// Mitsubishi GX Works2 project: SEMICON_SORTER_ENV   PLC: FX3U/FX3UC

PROGRAM MAIN
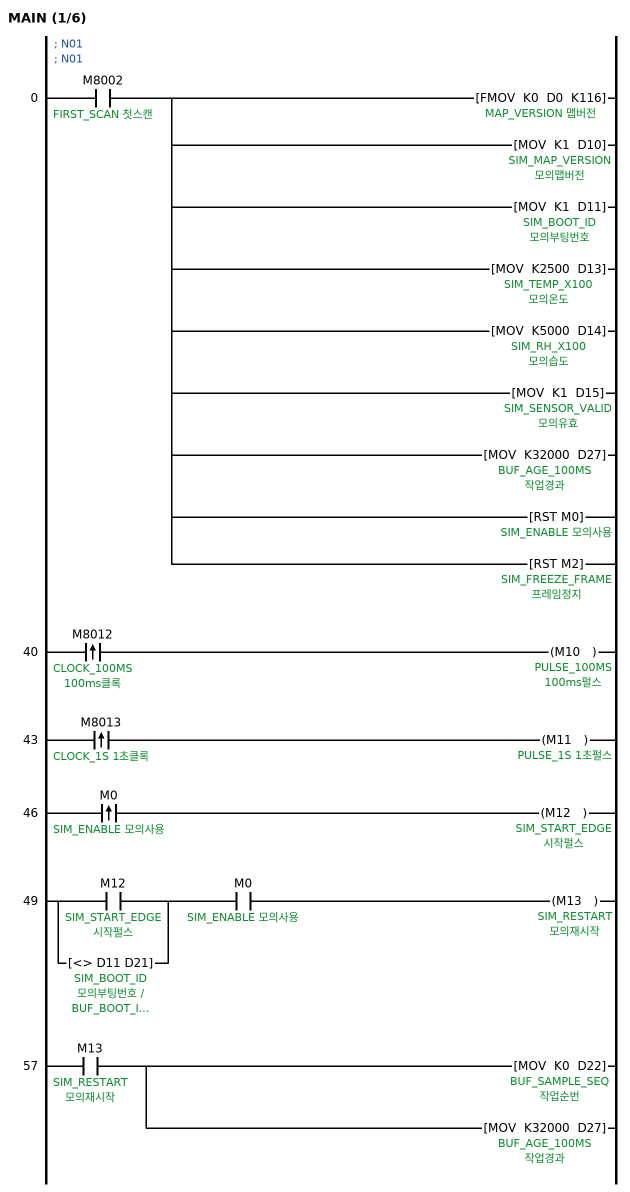
; 
; N01
; N01
0     LD      M8002  ; FIRST_SCAN 첫스캔
      FMOV    K0 D0 K116  ; MAP_VERSION 맵버전
      MOV     K1 D10  ; SIM_MAP_VERSION 모의맵버전
      MOV     K1 D11  ; SIM_BOOT_ID 모의부팅번호
      MOV     K2500 D13  ; SIM_TEMP_X100 모의온도
      MOV     K5000 D14  ; SIM_RH_X100 모의습도
      MOV     K1 D15  ; SIM_SENSOR_VALID 모의유효
      MOV     K32000 D27  ; BUF_AGE_100MS 작업경과
      RST     M0  ; SIM_ENABLE 모의사용
      RST     M2  ; SIM_FREEZE_FRAME 프레임정지
40    LDP     M8012  ; CLOCK_100MS 100ms클록
      OUT     M10  ; PULSE_100MS 100ms펄스
43    LDP     M8013  ; CLOCK_1S 1초클록
      OUT     M11  ; PULSE_1S 1초펄스
46    LDP     M0  ; SIM_ENABLE 모의사용
      OUT     M12  ; SIM_START_EDGE 시작펄스
49    LD      M12  ; SIM_START_EDGE 시작펄스
      OR<>    D11 D21  ; SIM_BOOT_ID 모의부팅번호 / BUF_BOOT_ID 작업부팅번호
      AND     M0  ; SIM_ENABLE 모의사용
      OUT     M13  ; SIM_RESTART 모의재시작
57    LD      M13  ; SIM_RESTART 모의재시작
      MOV     K0 D22  ; BUF_SAMPLE_SEQ 작업순번
      MOV     K32000 D27
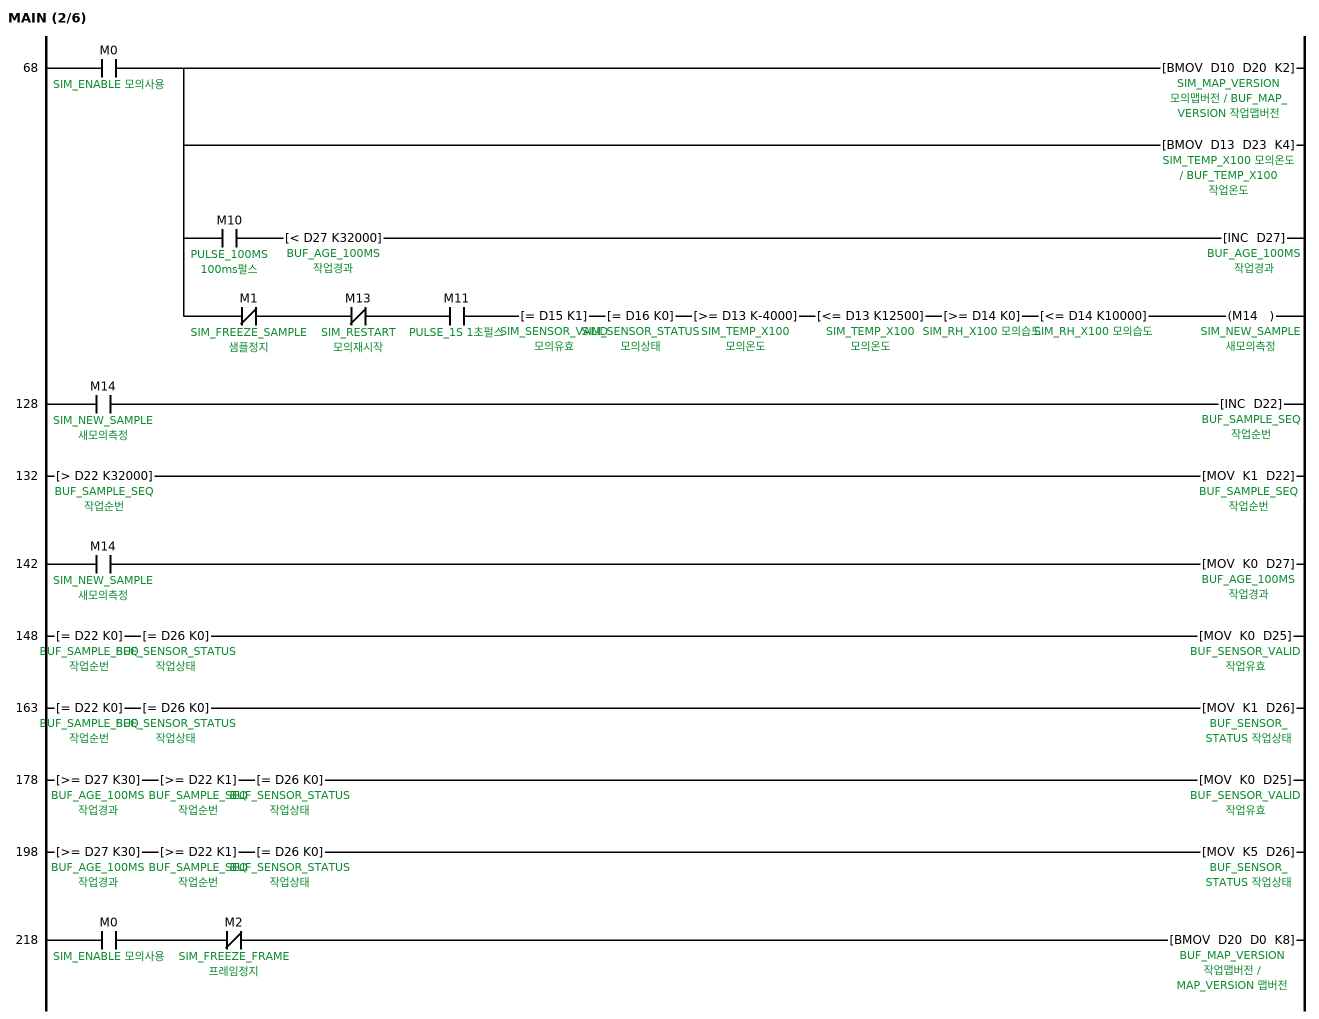
68    LD      M0  ; SIM_ENABLE 모의사용
      BMOV    D10 D20 K2  ; BUF_MAP_VERSION 작업맵버전
      BMOV    D13 D23 K4  ; BUF_TEMP_X100 작업온도
      MPS
      AND     M10  ; PULSE_100MS 100ms펄스
      AND<    D27 K32000  ; BUF_AGE_100MS 작업경과
      INC     D27
      MPP
      ANI     M1  ; SIM_FREEZE_SAMPLE 샘플정지
      ANI     M13  ; SIM_RESTART 모의재시작
      AND     M11  ; PULSE_1S 1초펄스
      AND=    D15 K1  ; SIM_SENSOR_VALID 모의유효
      AND=    D16 K0  ; SIM_SENSOR_STATUS 모의상태
      AND>=   D13 K-4000  ; SIM_TEMP_X100 모의온도
      AND<=   D13 K12500  ; SIM_TEMP_X100 모의온도
      AND>=   D14 K0  ; SIM_RH_X100 모의습도
      AND<=   D14 K10000  ; SIM_RH_X100 모의습도
      OUT     M14  ; SIM_NEW_SAMPLE 새모의측정
128   LD      M14  ; SIM_NEW_SAMPLE 새모의측정
      INC     D22
132   LD>     D22 K32000  ; BUF_SAMPLE_SEQ 작업순번
      MOV     K1 D22
142   LD      M14  ; SIM_NEW_SAMPLE 새모의측정
      MOV     K0 D27
148   LD=     D22 K0  ; BUF_SAMPLE_SEQ 작업순번
      AND=    D26 K0  ; BUF_SENSOR_STATUS 작업상태
      MOV     K0 D25  ; BUF_SENSOR_VALID 작업유효
163   LD=     D22 K0  ; BUF_SAMPLE_SEQ 작업순번
      AND=    D26 K0  ; BUF_SENSOR_STATUS 작업상태
      MOV     K1 D26
178   LD>=    D27 K30  ; BUF_AGE_100MS 작업경과
      AND>=   D22 K1  ; BUF_SAMPLE_SEQ 작업순번
      AND=    D26 K0  ; BUF_SENSOR_STATUS 작업상태
      MOV     K0 D25
198   LD>=    D27 K30  ; BUF_AGE_100MS 작업경과
      AND>=   D22 K1  ; BUF_SAMPLE_SEQ 작업순번
      AND=    D26 K0  ; BUF_SENSOR_STATUS 작업상태
      MOV     K5 D26
218   LD      M0  ; SIM_ENABLE 모의사용
      ANI     M2  ; SIM_FREEZE_FRAME 프레임정지
      BMOV    D20 D0 K8
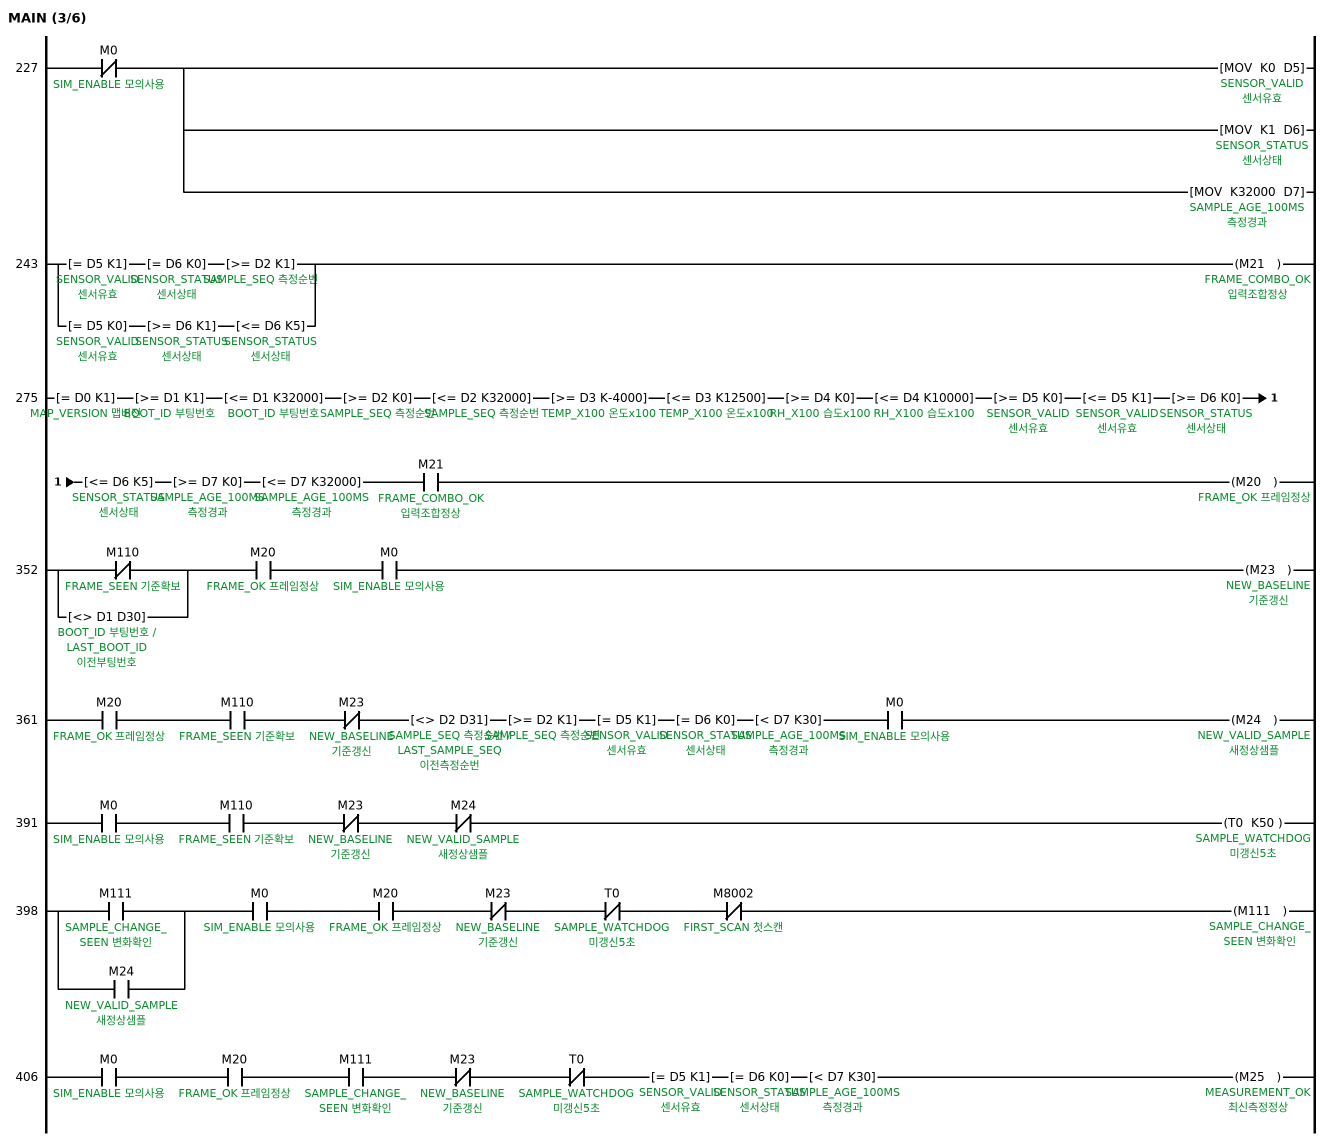
227   LDI     M0  ; SIM_ENABLE 모의사용
      MOV     K0 D5  ; SENSOR_VALID 센서유효
      MOV     K1 D6  ; SENSOR_STATUS 센서상태
      MOV     K32000 D7  ; SAMPLE_AGE_100MS 측정경과
243   LD=     D5 K1  ; SENSOR_VALID 센서유효
      AND=    D6 K0  ; SENSOR_STATUS 센서상태
      AND>=   D2 K1  ; SAMPLE_SEQ 측정순번
      LD=     D5 K0  ; SENSOR_VALID 센서유효
      AND>=   D6 K1  ; SENSOR_STATUS 센서상태
      AND<=   D6 K5  ; SENSOR_STATUS 센서상태
      ORB
      OUT     M21  ; FRAME_COMBO_OK 입력조합정상
275   LD=     D0 K1  ; MAP_VERSION 맵버전
      AND>=   D1 K1  ; BOOT_ID 부팅번호
      AND<=   D1 K32000  ; BOOT_ID 부팅번호
      AND>=   D2 K0  ; SAMPLE_SEQ 측정순번
      AND<=   D2 K32000  ; SAMPLE_SEQ 측정순번
      AND>=   D3 K-4000  ; TEMP_X100 온도x100
      AND<=   D3 K12500  ; TEMP_X100 온도x100
      AND>=   D4 K0  ; RH_X100 습도x100
      AND<=   D4 K10000  ; RH_X100 습도x100
      AND>=   D5 K0  ; SENSOR_VALID 센서유효
      AND<=   D5 K1  ; SENSOR_VALID 센서유효
      AND>=   D6 K0  ; SENSOR_STATUS 센서상태
      AND<=   D6 K5  ; SENSOR_STATUS 센서상태
      AND>=   D7 K0  ; SAMPLE_AGE_100MS 측정경과
      AND<=   D7 K32000  ; SAMPLE_AGE_100MS 측정경과
      AND     M21  ; FRAME_COMBO_OK 입력조합정상
      OUT     M20  ; FRAME_OK 프레임정상
352   LDI     M110  ; FRAME_SEEN 기준확보
      OR<>    D1 D30  ; BOOT_ID 부팅번호 / LAST_BOOT_ID 이전부팅번호
      AND     M20  ; FRAME_OK 프레임정상
      AND     M0  ; SIM_ENABLE 모의사용
      OUT     M23  ; NEW_BASELINE 기준갱신
361   LD      M20  ; FRAME_OK 프레임정상
      AND     M110  ; FRAME_SEEN 기준확보
      ANI     M23  ; NEW_BASELINE 기준갱신
      AND<>   D2 D31  ; SAMPLE_SEQ 측정순번 / LAST_SAMPLE_SEQ 이전측정순번
      AND>=   D2 K1  ; SAMPLE_SEQ 측정순번
      AND=    D5 K1  ; SENSOR_VALID 센서유효
      AND=    D6 K0  ; SENSOR_STATUS 센서상태
      AND<    D7 K30  ; SAMPLE_AGE_100MS 측정경과
      AND     M0  ; SIM_ENABLE 모의사용
      OUT     M24  ; NEW_VALID_SAMPLE 새정상샘플
391   LD      M0  ; SIM_ENABLE 모의사용
      AND     M110  ; FRAME_SEEN 기준확보
      ANI     M23  ; NEW_BASELINE 기준갱신
      ANI     M24  ; NEW_VALID_SAMPLE 새정상샘플
      OUT     T0 K50  ; SAMPLE_WATCHDOG 미갱신5초
398   LD      M111  ; SAMPLE_CHANGE_SEEN 변화확인
      OR      M24  ; NEW_VALID_SAMPLE 새정상샘플
      AND     M0  ; SIM_ENABLE 모의사용
      AND     M20  ; FRAME_OK 프레임정상
      ANI     M23  ; NEW_BASELINE 기준갱신
      ANI     T0  ; SAMPLE_WATCHDOG 미갱신5초
      ANI     M8002  ; FIRST_SCAN 첫스캔
      OUT     M111  ; SAMPLE_CHANGE_SEEN 변화확인
406   LD      M0  ; SIM_ENABLE 모의사용
      AND     M20  ; FRAME_OK 프레임정상
      AND     M111  ; SAMPLE_CHANGE_SEEN 변화확인
      ANI     M23  ; NEW_BASELINE 기준갱신
      ANI     T0  ; SAMPLE_WATCHDOG 미갱신5초
      AND=    D5 K1  ; SENSOR_VALID 센서유효
      AND=    D6 K0  ; SENSOR_STATUS 센서상태
      AND<    D7 K30  ; SAMPLE_AGE_100MS 측정경과
      OUT     M25  ; MEASUREMENT_OK 최신측정정상
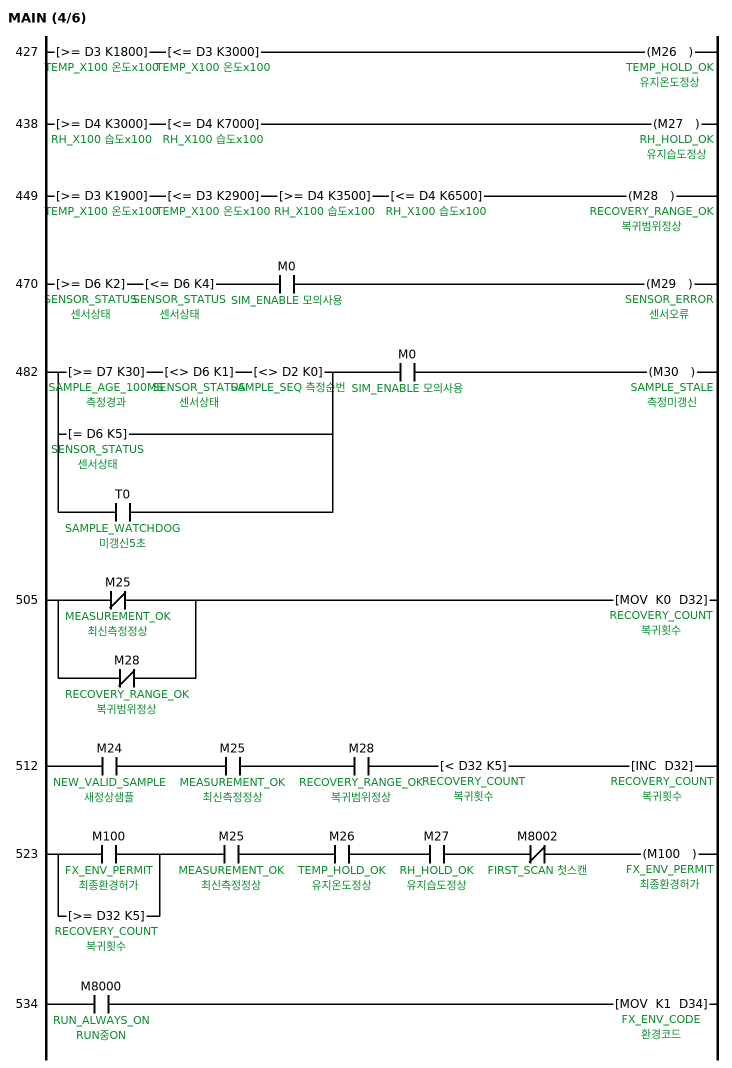
427   LD>=    D3 K1800  ; TEMP_X100 온도x100
      AND<=   D3 K3000  ; TEMP_X100 온도x100
      OUT     M26  ; TEMP_HOLD_OK 유지온도정상
438   LD>=    D4 K3000  ; RH_X100 습도x100
      AND<=   D4 K7000  ; RH_X100 습도x100
      OUT     M27  ; RH_HOLD_OK 유지습도정상
449   LD>=    D3 K1900  ; TEMP_X100 온도x100
      AND<=   D3 K2900  ; TEMP_X100 온도x100
      AND>=   D4 K3500  ; RH_X100 습도x100
      AND<=   D4 K6500  ; RH_X100 습도x100
      OUT     M28  ; RECOVERY_RANGE_OK 복귀범위정상
470   LD>=    D6 K2  ; SENSOR_STATUS 센서상태
      AND<=   D6 K4  ; SENSOR_STATUS 센서상태
      AND     M0  ; SIM_ENABLE 모의사용
      OUT     M29  ; SENSOR_ERROR 센서오류
482   LD>=    D7 K30  ; SAMPLE_AGE_100MS 측정경과
      AND<>   D6 K1  ; SENSOR_STATUS 센서상태
      AND<>   D2 K0  ; SAMPLE_SEQ 측정순번
      OR=     D6 K5  ; SENSOR_STATUS 센서상태
      OR      T0  ; SAMPLE_WATCHDOG 미갱신5초
      AND     M0  ; SIM_ENABLE 모의사용
      OUT     M30  ; SAMPLE_STALE 측정미갱신
505   LDI     M25  ; MEASUREMENT_OK 최신측정정상
      ORI     M28  ; RECOVERY_RANGE_OK 복귀범위정상
      MOV     K0 D32  ; RECOVERY_COUNT 복귀횟수
512   LD      M24  ; NEW_VALID_SAMPLE 새정상샘플
      AND     M25  ; MEASUREMENT_OK 최신측정정상
      AND     M28  ; RECOVERY_RANGE_OK 복귀범위정상
      AND<    D32 K5  ; RECOVERY_COUNT 복귀횟수
      INC     D32
523   LD      M100  ; FX_ENV_PERMIT 최종환경허가
      OR>=    D32 K5  ; RECOVERY_COUNT 복귀횟수
      AND     M25  ; MEASUREMENT_OK 최신측정정상
      AND     M26  ; TEMP_HOLD_OK 유지온도정상
      AND     M27  ; RH_HOLD_OK 유지습도정상
      ANI     M8002  ; FIRST_SCAN 첫스캔
      OUT     M100  ; FX_ENV_PERMIT 최종환경허가
534   LD      M8000  ; RUN_ALWAYS_ON RUN중ON
      MOV     K1 D34  ; FX_ENV_CODE 환경코드
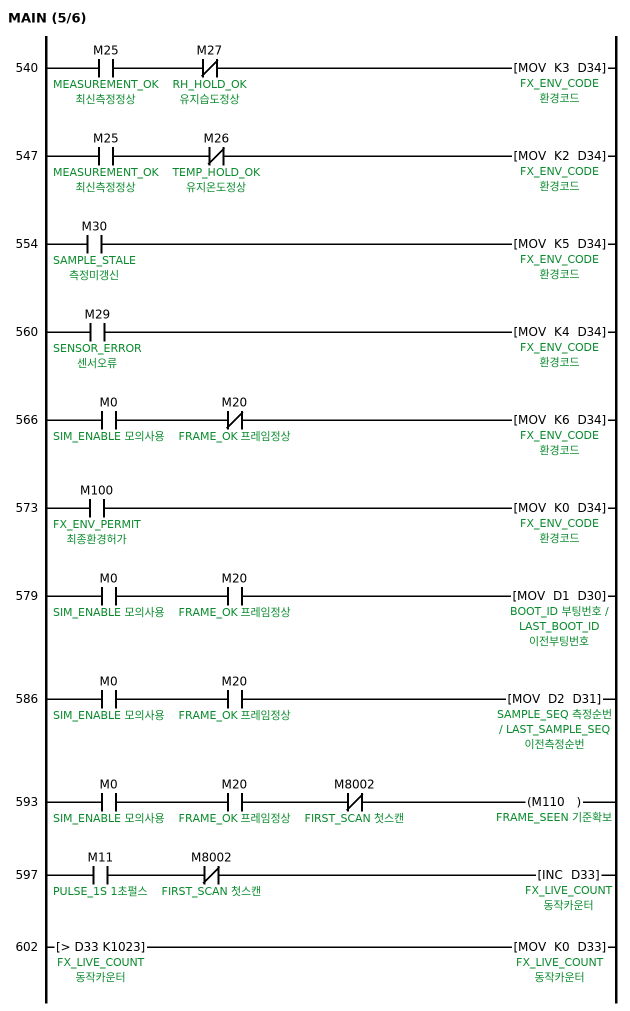
540   LD      M25  ; MEASUREMENT_OK 최신측정정상
      ANI     M27  ; RH_HOLD_OK 유지습도정상
      MOV     K3 D34
547   LD      M25  ; MEASUREMENT_OK 최신측정정상
      ANI     M26  ; TEMP_HOLD_OK 유지온도정상
      MOV     K2 D34
554   LD      M30  ; SAMPLE_STALE 측정미갱신
      MOV     K5 D34
560   LD      M29  ; SENSOR_ERROR 센서오류
      MOV     K4 D34
566   LD      M0  ; SIM_ENABLE 모의사용
      ANI     M20  ; FRAME_OK 프레임정상
      MOV     K6 D34
573   LD      M100  ; FX_ENV_PERMIT 최종환경허가
      MOV     K0 D34
579   LD      M0  ; SIM_ENABLE 모의사용
      AND     M20  ; FRAME_OK 프레임정상
      MOV     D1 D30
586   LD      M0  ; SIM_ENABLE 모의사용
      AND     M20  ; FRAME_OK 프레임정상
      MOV     D2 D31
593   LD      M0  ; SIM_ENABLE 모의사용
      AND     M20  ; FRAME_OK 프레임정상
      ANI     M8002  ; FIRST_SCAN 첫스캔
      OUT     M110  ; FRAME_SEEN 기준확보
597   LD      M11  ; PULSE_1S 1초펄스
      ANI     M8002  ; FIRST_SCAN 첫스캔
      INC     D33  ; FX_LIVE_COUNT 동작카운터
602   LD>     D33 K1023  ; FX_LIVE_COUNT 동작카운터
      MOV     K0 D33
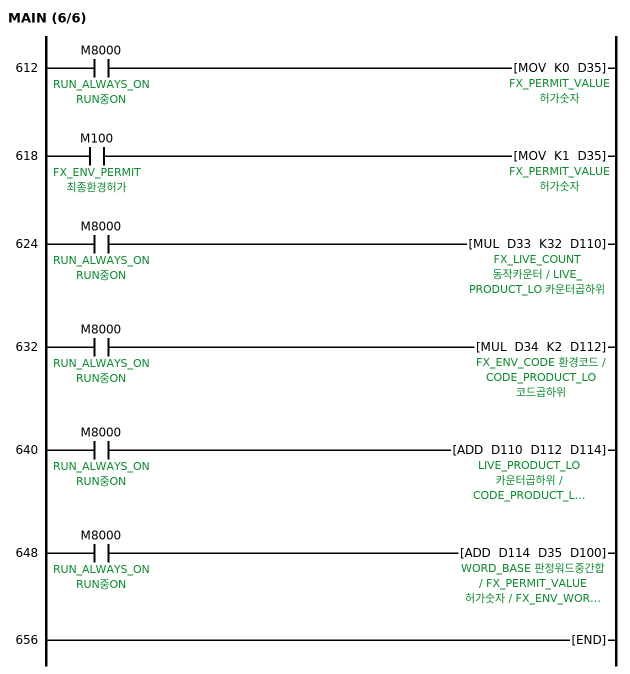
612   LD      M8000  ; RUN_ALWAYS_ON RUN중ON
      MOV     K0 D35  ; FX_PERMIT_VALUE 허가숫자
618   LD      M100  ; FX_ENV_PERMIT 최종환경허가
      MOV     K1 D35
624   LD      M8000  ; RUN_ALWAYS_ON RUN중ON
      MUL     D33 K32 D110  ; LIVE_PRODUCT_LO 카운터곱하위
632   LD      M8000  ; RUN_ALWAYS_ON RUN중ON
      MUL     D34 K2 D112  ; CODE_PRODUCT_LO 코드곱하위
640   LD      M8000  ; RUN_ALWAYS_ON RUN중ON
      ADD     D110 D112 D114  ; WORD_BASE 판정워드중간합
648   LD      M8000  ; RUN_ALWAYS_ON RUN중ON
      ADD     D114 D35 D100  ; FX_ENV_WORD 최종판정워드
656   END
END_PROGRAM

// device comments not shown above
D24  ; BUF_RH_X100 작업습도
D111  ; LIVE_PRODUCT_HI 카운터곱상위
D113  ; CODE_PRODUCT_HI 코드곱상위
D115  ; RESERVED 예약미사용
